// TIA Portal V21 export
// export: Created 2026-11-10T19:11:35.9319997Z, ExportSetting WithDefaults, DisplayName Totally Integrated Automation Portal, DisplayVersion V21 Update 3, DisplayName STEP 7 Professional, DisplayVersion V21 Update 3, DisplayName STEP 7 Safety, DisplayVersion V21, DisplayName Tech WebApplication, DisplayVersion V21, DisplayName WinCC Basic/Comfort/Advanced, DisplayVersion V21 Update 3, DisplayName WinCC Unified, DisplayVersion V21 Update 3
DATA_BLOCK "DB_GETIO_PART"   // DB19
// stored: AutoNumber true, DBAccessibleFromOPCUA true, DBAccessibleFromWebserver true, InstanceOfName GETIO_PART, OfSystemLibElement GETIO_PART, OfSystemLibVersion 1.2
"GETIO_PART"
   // VAR_INPUT
   //    ID : HW_SUBMODULE;
   //    OFFSET : Int;
   //    LEN : Int;
   // END_VAR
   // VAR_OUTPUT
   //    STATUS : DWord;
   //    ERROR : Bool;
   // END_VAR
   // VAR_IN_OUT
   //    INPUTS : Variant;
   // END_VAR
BEGIN
END_DATA_BLOCK
